Fanuc KAREL source: kx00031.KL

-- PROVISIONAL review KL for V770-1; original PC SHA256 f70c0f127969fee2eb76dcbb31f58be78b37eeb6fecb9fdc011aa7cce3c25799
-- Incomplete behavior may be omitted. Consult companion uncertainty JSON. Do not deploy.
PROGRAM KX00031
%NOLOCKGROUP
VAR
  I : INTEGER
  J : INTEGER
  B : BOOLEAN
  F : FILE
  S : STRING[80]
-- UNRESOLVED_DECL P type=000102
BEGIN
  -- UNRESOLVED_PC offsets 5-12; opcodes 9D,23
  -- UNRESOLVED_PC offsets 17-21; opcodes 7F
END KX00031
